// TIA Portal V21 export
// export: Created 2026-10-24T00:49:22.4780738Z, ExportSetting WithDefaults, DisplayName Totally Integrated Automation Portal, DisplayVersion V21 Update 1, DisplayName SINAMICS Startdrive Advanced, DisplayVersion V21 HF2, DisplayName SINAMICS Startdrive G110M, G120, G120C, G120D, G120P, G115D, DisplayVersion V21 HF2, DisplayName SINAMICS Startdrive G130, G150, S120, S150, G200, G220, S200, S210, S220, Innomotics MVD, DisplayVersion V21 HF2, DisplayName STEP 7 Professional, DisplayVersion V21 Update 1, DisplayName STEP 7 Safety, DisplayVersion V21, DisplayName Tech WebApplication, DisplayVersion V21, DisplayName WinCC Basic/Comfort/Advanced, DisplayVersion V21 Update 1, DisplayName WinCC Unified, DisplayVersion V21 Update 1
VAR_GLOBAL   // PLC tag table "Tags_Memory"
   HelperBit AT %M10.0 : Bool;   // Hilfsmerker / Helper bit
   PulseBit AT %M10.1 : Bool;   // Impulsmerker / Pulse bit
   StatusMemoryWord AT %MW12 : Word;   // Statuswort / Status word
   PieceCountMemory AT %MW14 : Int;   // Stückzahl / Piece count
   ServiceWord AT %MW16 : Word;   // Servicewort, nicht von HMI erreichbar / Service word, not accessible from HMI   {ExternalAccessible false, ExternalVisible false, ExternalWritable false}
END_VAR
VAR_GLOBAL CONSTANT   // user constants
   MAXIMUM_PIECES : Int := 1000;   // Maximale Stückzahl pro Charge / Maximum pieces per batch
   NOMINAL_FLOW : Real := 12.5;   // Nenndurchfluss in l/min / Nominal flow in l/min
   FILL_TIMEOUT : Time := T#30s;   // Füllzeitüberschreitung / Filling timeout
END_VAR
